(* IEC 61131-3 sources: plc-vscode/tests/st/all/trust-platform/examples/OSCAT/district_pump_network_proxy_mediator/non-oop/src, 3 files *)

(* ---- Main.st ---- *)
FUNCTION_BLOCK ClassicDistrictPumpNetwork
VAR
    TotalDemandM3HValue : REAL;
    PumpSpeedPctValue : REAL;
    RemoteStaleCountValue : INT;
    ClassAAlarmValue : BOOL;
END_VAR

METHOD PUBLIC Update : REAL
VAR_INPUT
    LocalDemandM3H : REAL;
    NorthDemandM3H : REAL;
    NorthQualityGood : BOOL;
    NorthAgeSeconds : INT;
    EastDemandM3H : REAL;
    EastQualityGood : BOOL;
    EastAgeSeconds : INT;
    SuctionHealthy : BOOL;
END_VAR
TotalDemandM3HValue := LocalDemandM3H;
RemoteStaleCountValue := INT#0;

IF NorthQualityGood AND (NorthAgeSeconds <= INT#30) THEN
    TotalDemandM3HValue := TotalDemandM3HValue + NorthDemandM3H;
ELSE
    RemoteStaleCountValue := RemoteStaleCountValue + INT#1;
END_IF;

IF EastQualityGood AND (EastAgeSeconds <= INT#30) THEN
    TotalDemandM3HValue := TotalDemandM3HValue + EastDemandM3H;
ELSE
    RemoteStaleCountValue := RemoteStaleCountValue + INT#1;
END_IF;

ClassAAlarmValue := NOT SuctionHealthy;
IF ClassAAlarmValue THEN
    PumpSpeedPctValue := REAL#0.0;
ELSE
    PumpSpeedPctValue := LIMIT(REAL#0.0, TotalDemandM3HValue * REAL#2.0, REAL#100.0);
END_IF;
Update := PumpSpeedPctValue;
END_METHOD

PUBLIC PROPERTY TotalDemandM3H : REAL
GET
    TotalDemandM3H := TotalDemandM3HValue;
END_GET
END_PROPERTY

PUBLIC PROPERTY RemoteStaleCount : INT
GET
    RemoteStaleCount := RemoteStaleCountValue;
END_GET
END_PROPERTY

PUBLIC PROPERTY ClassAAlarm : BOOL
GET
    ClassAAlarm := ClassAAlarmValue;
END_GET
END_PROPERTY
END_FUNCTION_BLOCK

PROGRAM Main
VAR
    Network : ClassicDistrictPumpNetwork;
    LocalDemandRaw : INT;
    NorthDemandRaw : INT;
    EastDemandRaw : INT;
    NorthAgeSeconds : INT;
    EastAgeSeconds : INT;
    NorthQualityGood : BOOL;
    EastQualityGood : BOOL;
    SuctionHealthy : BOOL;
    PumpSpeedRaw : INT;
    StaleAlarmOut : BOOL;
END_VAR
Network.Update(LocalDemandM3H := INT_TO_REAL(LocalDemandRaw), NorthDemandM3H := INT_TO_REAL(NorthDemandRaw), NorthQualityGood := NorthQualityGood, NorthAgeSeconds := NorthAgeSeconds, EastDemandM3H := INT_TO_REAL(EastDemandRaw), EastQualityGood := EastQualityGood, EastAgeSeconds := EastAgeSeconds, SuctionHealthy := SuctionHealthy);
PumpSpeedRaw := REAL_TO_INT(Network.Update(LocalDemandM3H := INT_TO_REAL(LocalDemandRaw), NorthDemandM3H := INT_TO_REAL(NorthDemandRaw), NorthQualityGood := NorthQualityGood, NorthAgeSeconds := NorthAgeSeconds, EastDemandM3H := INT_TO_REAL(EastDemandRaw), EastQualityGood := EastQualityGood, EastAgeSeconds := EastAgeSeconds, SuctionHealthy := SuctionHealthy));
StaleAlarmOut := Network.RemoteStaleCount > INT#0;
END_PROGRAM

(* ---- Configuration.st ---- *)
CONFIGURATION DistrictPumpNetworkProxyMediatorClassicConfiguration
RESOURCE Cpu0 ON PLC
    TASK MainTask (INTERVAL := T#100ms, PRIORITY := 1);
    PROGRAM Network WITH MainTask : Main;
END_RESOURCE
VAR_CONFIG
    Network.LocalDemandRaw AT %IW0 : INT;
    Network.NorthDemandRaw AT %IW2 : INT;
    Network.EastDemandRaw AT %IW4 : INT;
    Network.NorthAgeSeconds AT %IW6 : INT;
    Network.EastAgeSeconds AT %IW8 : INT;
    Network.NorthQualityGood AT %IX0.0 : BOOL;
    Network.EastQualityGood AT %IX0.1 : BOOL;
    Network.SuctionHealthy AT %IX0.2 : BOOL;
    Network.PumpSpeedRaw AT %QW0 : INT;
    Network.StaleAlarmOut AT %QX0.0 : BOOL;
END_VAR
END_CONFIGURATION

(* ---- Tests.st ---- *)
TEST_PROGRAM ClassicDistrictBalancesHealthyDemand
VAR
    Network : ClassicDistrictPumpNetwork;
END_VAR

ASSERT_EQUAL(EXPECTED := REAL#90.0, ACTUAL := Network.Update(LocalDemandM3H := REAL#20.0, NorthDemandM3H := REAL#15.0, NorthQualityGood := TRUE, NorthAgeSeconds := INT#5, EastDemandM3H := REAL#10.0, EastQualityGood := TRUE, EastAgeSeconds := INT#5, SuctionHealthy := TRUE));
ASSERT_EQUAL(EXPECTED := REAL#45.0, ACTUAL := Network.TotalDemandM3H);
END_TEST_PROGRAM

TEST_PROGRAM ClassicDistrictDropsStaleDemand
VAR
    Network : ClassicDistrictPumpNetwork;
END_VAR

ASSERT_EQUAL(EXPECTED := REAL#40.0, ACTUAL := Network.Update(LocalDemandM3H := REAL#20.0, NorthDemandM3H := REAL#15.0, NorthQualityGood := TRUE, NorthAgeSeconds := INT#45, EastDemandM3H := REAL#10.0, EastQualityGood := FALSE, EastAgeSeconds := INT#5, SuctionHealthy := TRUE));
ASSERT_EQUAL(EXPECTED := INT#2, ACTUAL := Network.RemoteStaleCount);
END_TEST_PROGRAM
